(* Logix 5000 project; controller R400_500_XLS vendor 1 type 14 code 216 rev 31.11; software revision 31.01; part 16 of 32 *)
(* tags used below, declared in another part *)
   CycleModifBuffer : UDT_CYCLE;
   DRYING : DINT;   // Drying id number
   DRYING_HEAT_SENSITIVE_SEL : DINT;   // Drying heat sensitive
   DRYING_MODE_SEL : DINT;   // Drying mode selector index
   DRYING_TEMP_C_SEL : DINT;   // Drying temperature index
   DRYING_TEMP_F_SEL : DINT;   // Drying temperature index
   DRYING_TIME_MIN_NUM : DINT;   // Drying time (minutes) numeric input index
   DRYING_TIME_SEC_NUM : DINT;   // Drying time (seconds) numeric input index
   FC83_DryHeatSensitive : DINT;   // Drying is heat sensitive?
   FC83_DryTemp : DINT;   // Drying temperature (hi/low)
   FC83_FRinse_Drained : DINT;   // Drained final rinse flag
   FC83_FRinse_Heated : DINT;   // Heated final rinse flag
   FC83_FRinse_Recirculated : DINT;   // Recirculated final rinse flag
   FC83_ONS : SINT;
   FRINSE_COND_SET_POINT_NUM : DINT;   // Final rinse conductivity set point numeric input index
   FRINSE_DRAIN_SEL : DINT;   // Final rinse drained selector's index
   FRINSE_HEATING_SEL : DINT;   // Final rinse heating selector's index
   FRINSE_MIN_NUMBER_NUM : DINT;   // Final rinse minimum number of final rinse numeric input index
   FRINSE_NUMBER_NUM : DINT;   // Final rinse number of final rinse numeric input index
   FRINSE_RECIRC_SEL : DINT;   // Final rinse recirculated selector's index
   FRINSE_TIME_MIN_NUM : DINT;   // Final rinse time (minutes) numeric input index
   FRINSE_TIME_SEC_NUM : DINT;   // Final rinse time (seconds) numeric input index
   FRINSE_TYPE_SEL : DINT;   // Final rinse type selector's index
   M : DINT[5];   // Memory Bits
   MaxTrtTempSp : REAL;
   NON_RECIRCULATED_FINAL_RINSE_MINUTES : DINT;   // Number of minutes for the non recirculated final rinse
   NON_RECIRCULATED_FINAL_RINSE_SECONDS : DINT;   // Number of seconds for the non recirculated final rinse
   Rinse_Select : BOOL;
   RinseIndex : SINT;
   Second_Inj_conc : BOOL;
   WashIndex : SINT;
   cfgRinseHeated : SINT;
   cfgRinseMin : SINT;
   cfgRinseSec : SINT;
   CfgRinseTempSp : REAL;
   cfgRinseWport : SINT;
   CfgWshInjRateImperial : REAL;   // Wash Injection Rate - Oz / Gal
   CfgWshInjRateMetric : REAL;   // Wash Injection Rate - mL / L
   ChemConcUnit : BOOL;   // 0 = mL/L; 1 = oz/gal
   Msg_TempSp : SINT;   // HMI Information Message tag
   NumInput : UDT_NUMERIC_INPUT[65];   // Numeric input
   NumInputReal : UDT_NUMERIC_INPUT_REAL[17];
   Screen_Ctrl : DINT;   // PLC Screen Request
   Selector : UDT_SELECTOR[25];   // Piloted list selector
   TempUnit : BOOL;   // Temperature Units 0= Celcius 1 = Farhenheit
   Tpb : DINT[11];
   TpbImage : DINT[11];
   udtFRHeatingSel : UDT_SELECTOR;
   udtFRLastRinseDrained : UDT_SELECTOR;
   udtFRRecirculation : UDT_SELECTOR;
   udtFRType : UDT_SELECTOR;
   Unit : Hrdwre;   // Unit Configuration
(* MainProgram, continued *)

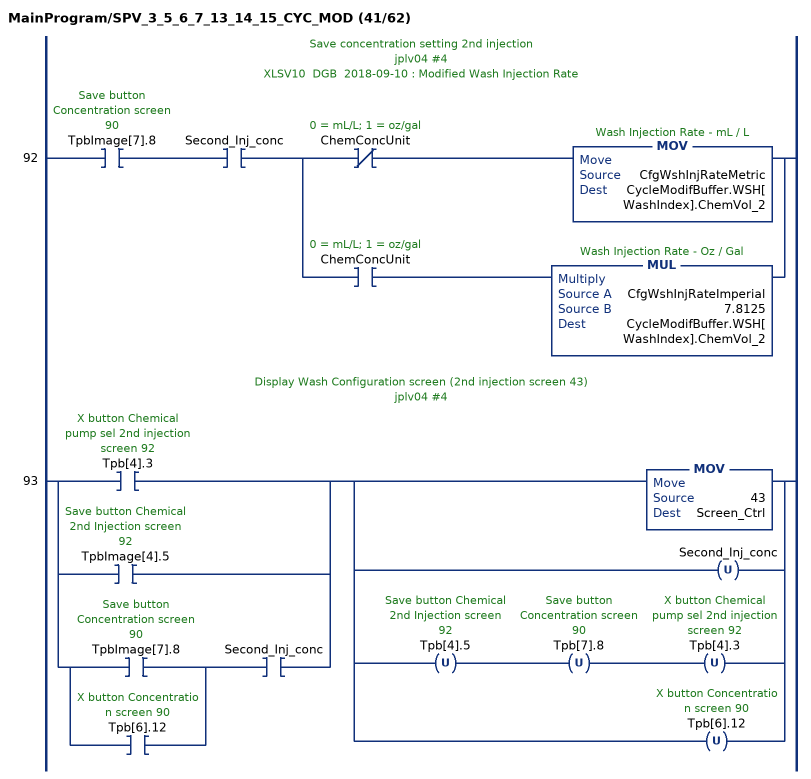
   [picture p292: MainProgram/SPV_3_5_6_7_13_14_15_CYC_MOD rungs 92-93]
   // Save concentration setting 2nd injection
   // jplv04 #4
   // XLSV10  DGB  2018-09-10 : Modified Wash Injection Rate
   92: XIC(TpbImage[7].8)XIC(Second_Inj_conc)[XIO(ChemConcUnit) MOV(CfgWshInjRateMetric,CycleModifBuffer.WSH[WashIndex].ChemVol_2) ,XIC(ChemConcUnit) MUL(CfgWshInjRateImperial,7.8125,CycleModifBuffer.WSH[WashIndex].ChemVol_2) ];
   // Display Wash Configuration screen (2nd injection screen 43)
   // jplv04 #4
   93: [XIC(Tpb[4].3) ,XIC(TpbImage[4].5) ,[XIC(TpbImage[7].8) ,XIC(Tpb[6].12) ] XIC(Second_Inj_conc) ][MOV(43,Screen_Ctrl) ,OTU(Second_Inj_conc) ,OTU(Tpb[4].5) OTU(Tpb[7].8) OTU(Tpb[4].3) ,OTU(Tpb[6].12) ];
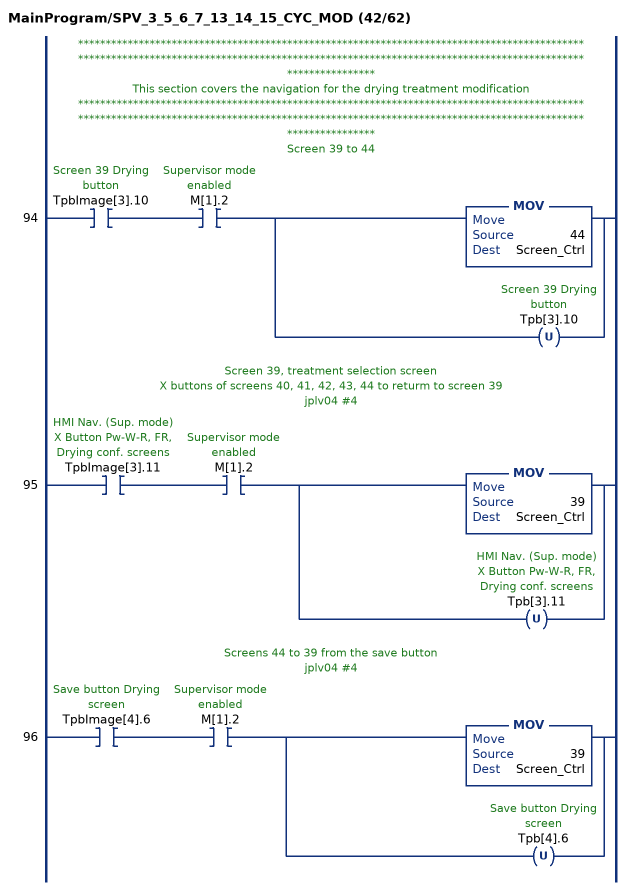
   // ********************************************************************************************************************************************************************************************************
   // This section covers the navigation for the drying treatment modification
   // ********************************************************************************************************************************************************************************************************
   // Screen 39 to 44
   94: XIC(TpbImage[3].10)XIC(M[1].2)[MOV(44,Screen_Ctrl) ,OTU(Tpb[3].10) ];
   // Screen 39, treatment selection screen
   // X buttons of screens 40, 41, 42, 43, 44 to returm to screen 39
   // jplv04 #4
   95: XIC(TpbImage[3].11)XIC(M[1].2)[MOV(39,Screen_Ctrl) ,OTU(Tpb[3].11) ];
   // Screens 44 to 39 from the save button
   // jplv04 #4
   96: XIC(TpbImage[4].6)XIC(M[1].2)[MOV(39,Screen_Ctrl) ,OTU(Tpb[4].6) ];
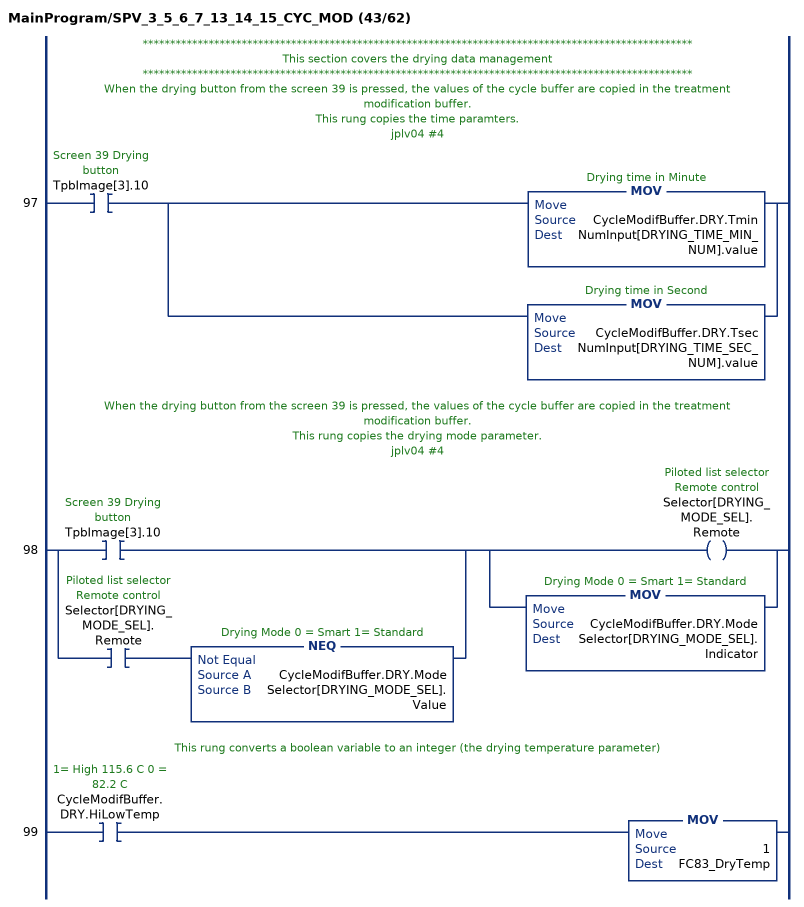
   // ****************************************************************************************************
   // This section covers the drying data management
   // ****************************************************************************************************
   // When the drying button from the screen 39 is pressed, the values of the cycle buffer are copied in the treatment modification buffer.
   // This rung copies the time paramters.
   // jplv04 #4
   97: XIC(TpbImage[3].10)[MOV(CycleModifBuffer.DRY.Tmin,NumInput[DRYING_TIME_MIN_NUM].value) ,MOV(CycleModifBuffer.DRY.Tsec,NumInput[DRYING_TIME_SEC_NUM].value) ];
   // When the drying button from the screen 39 is pressed, the values of the cycle buffer are copied in the treatment modification buffer.
   // This rung copies the drying mode parameter.
   // jplv04 #4
   98: [XIC(TpbImage[3].10) ,XIC(Selector[DRYING_MODE_SEL].Remote) NEQ(CycleModifBuffer.DRY.Mode,Selector[DRYING_MODE_SEL].Value) ][OTE(Selector[DRYING_MODE_SEL].Remote) ,MOV(CycleModifBuffer.DRY.Mode,Selector[DRYING_MODE_SEL].Indicator) ];
   // This rung converts a boolean variable to an integer (the drying temperature parameter)
   99: XIC(CycleModifBuffer.DRY.HiLowTemp)MOV(1,FC83_DryTemp);
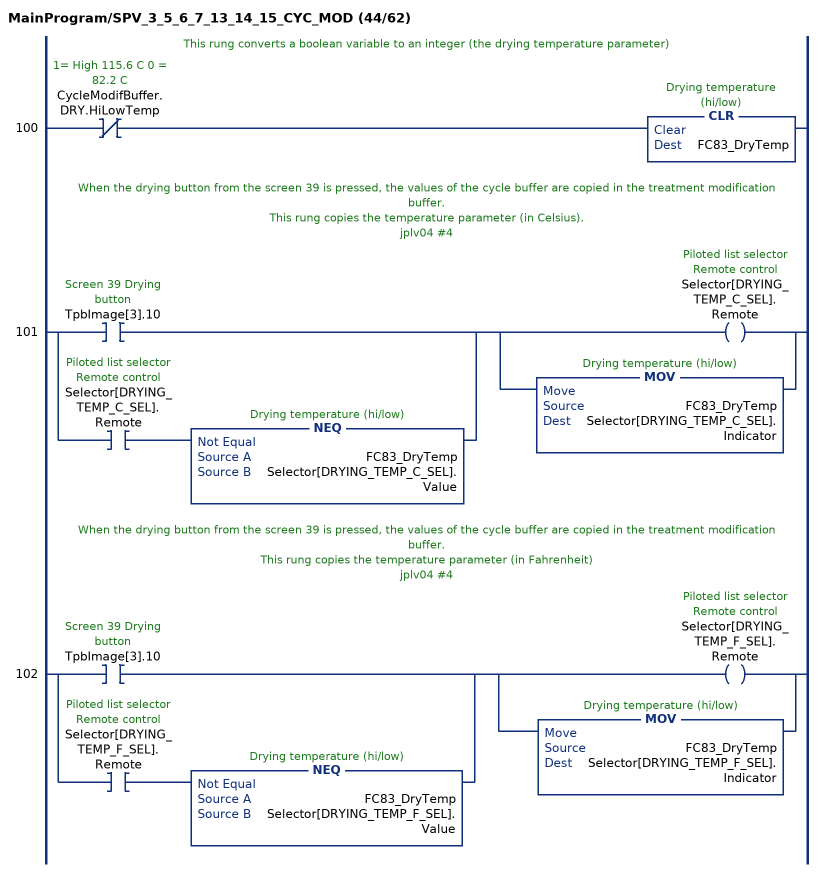
   // This rung converts a boolean variable to an integer (the drying temperature parameter)
   100: XIO(CycleModifBuffer.DRY.HiLowTemp)CLR(FC83_DryTemp);
   // When the drying button from the screen 39 is pressed, the values of the cycle buffer are copied in the treatment modification buffer.
   // This rung copies the temperature parameter (in Celsius).
   // jplv04 #4
   101: [XIC(TpbImage[3].10) ,XIC(Selector[DRYING_TEMP_C_SEL].Remote) NEQ(FC83_DryTemp,Selector[DRYING_TEMP_C_SEL].Value) ][OTE(Selector[DRYING_TEMP_C_SEL].Remote) ,MOV(FC83_DryTemp,Selector[DRYING_TEMP_C_SEL].Indicator) ];
   // When the drying button from the screen 39 is pressed, the values of the cycle buffer are copied in the treatment modification buffer.
   // This rung copies the temperature parameter (in Fahrenheit)
   // jplv04 #4
   102: [XIC(TpbImage[3].10) ,XIC(Selector[DRYING_TEMP_F_SEL].Remote) NEQ(FC83_DryTemp,Selector[DRYING_TEMP_F_SEL].Value) ][OTE(Selector[DRYING_TEMP_F_SEL].Remote) ,MOV(FC83_DryTemp,Selector[DRYING_TEMP_F_SEL].Indicator) ];
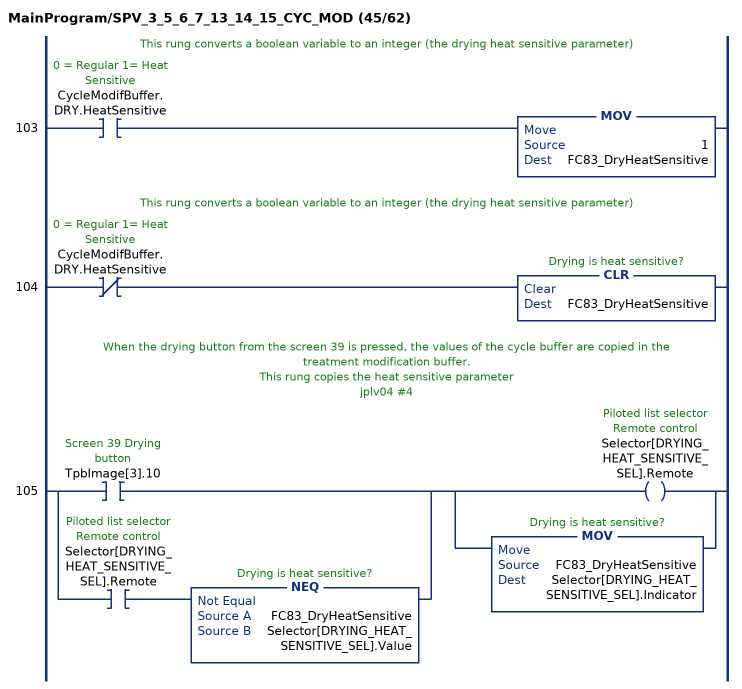
   // This rung converts a boolean variable to an integer (the drying heat sensitive parameter)
   103: XIC(CycleModifBuffer.DRY.HeatSensitive)MOV(1,FC83_DryHeatSensitive);
   // This rung converts a boolean variable to an integer (the drying heat sensitive parameter)
   104: XIO(CycleModifBuffer.DRY.HeatSensitive)CLR(FC83_DryHeatSensitive);
   // When the drying button from the screen 39 is pressed, the values of the cycle buffer are copied in the treatment modification buffer.
   // This rung copies the heat sensitive parameter
   // jplv04 #4
   105: [XIC(TpbImage[3].10) ,XIC(Selector[DRYING_HEAT_SENSITIVE_SEL].Remote) NEQ(FC83_DryHeatSensitive,Selector[DRYING_HEAT_SENSITIVE_SEL].Value) ][OTE(Selector[DRYING_HEAT_SENSITIVE_SEL].Remote) ,MOV(FC83_DryHeatSensitive,Selector[DRYING_HEAT_SENSITIVE_SEL].Indicator) ];
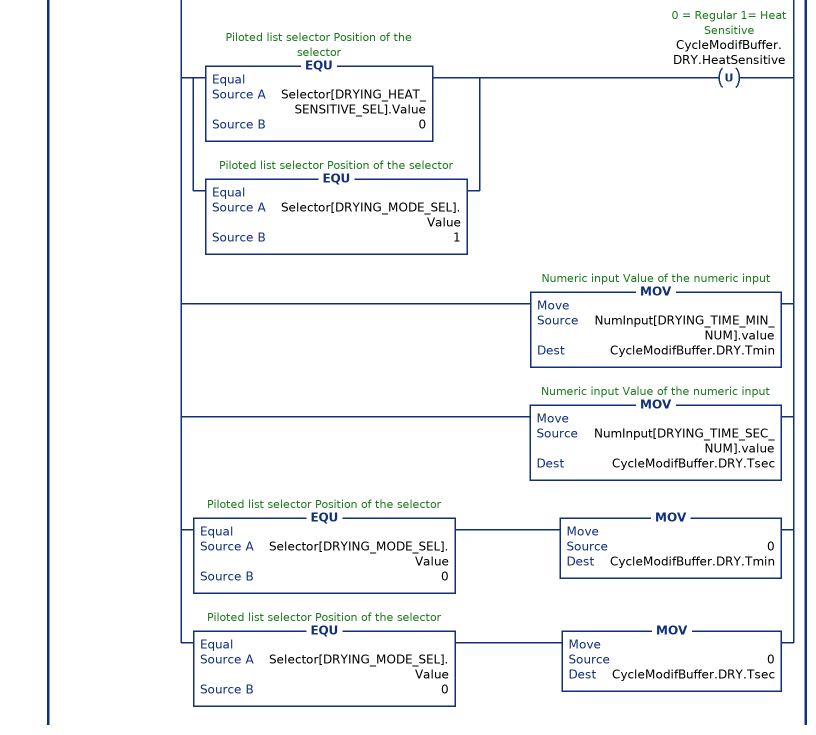
   // When the save button is pressed, the values are copied from the drying modification buffer to the cycle modification buffer
   // jplv04 #4
   106: XIC(TpbImage[4].6)[MOV(Selector[DRYING_MODE_SEL].Value,CycleModifBuffer.DRY.Mode) ,[XIO(TempUnit) EQU(Selector[DRYING_TEMP_C_SEL].Value,1) ,XIC(TempUnit) EQU(Selector[DRYING_TEMP_F_SEL].Value,1) ] OTL(CycleModifBuffer.DRY.HiLowTemp) ,[XIC(TempUnit) EQU(Selector[DRYING_TEMP_F_SEL].Value,0) ,XIO(TempUnit) EQU(Selector[DRYING_TEMP_C_SEL].Value,0) ,EQU(Selector[DRYING_MODE_SEL].Value,0) ] OTU(CycleModifBuffer.DRY.HiLowTemp) ,EQU(Selector[DRYING_HEAT_SENSITIVE_SEL].Value,1) OTL(CycleModifBuffer.DRY.HeatSensitive) ,[EQU(Selector[DRYING_HEAT_SENSITIVE_SEL].Value,0) ,EQU(Selector[DRYING_MODE_SEL].Value,1) ] OTU(CycleModifBuffer.DRY.HeatSensitive) ,MOV(NumInput[DRYING_TIME_MIN_NUM].value,CycleModifBuffer.DRY.Tmin) ,MOV(NumInput[DRYING_TIME_SEC_NUM].value,CycleModifBuffer.DRY.Tsec) ,EQU(Selector[DRYING_MODE_SEL].Value,0) MOV(0,CycleModifBuffer.DRY.Tmin) ,EQU(Selector[DRYING_MODE_SEL].Value,0) MOV(0,CycleModifBuffer.DRY.Tsec) ];
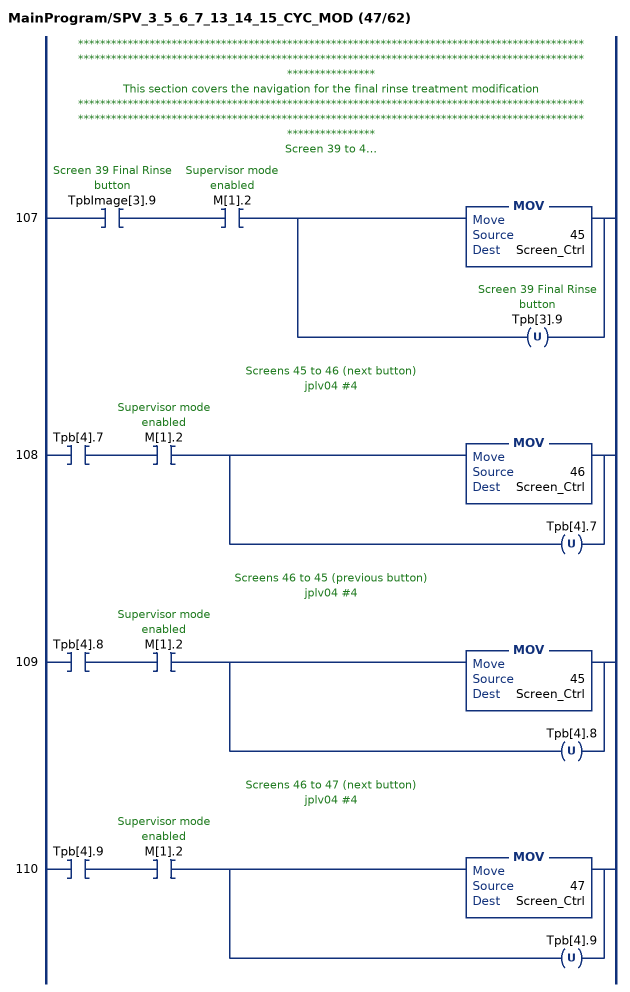
   // ********************************************************************************************************************************************************************************************************
   // This section covers the navigation for the final rinse treatment modification
   // ********************************************************************************************************************************************************************************************************
   // Screen 39 to 45
   // jplv04 #4
   107: XIC(TpbImage[3].9)XIC(M[1].2)[MOV(45,Screen_Ctrl) ,OTU(Tpb[3].9) ];
   // Screens 45 to 46 (next button)
   // jplv04 #4
   108: XIC(Tpb[4].7)XIC(M[1].2)[MOV(46,Screen_Ctrl) ,OTU(Tpb[4].7) ];
   // Screens 46 to 45 (previous button)
   // jplv04 #4
   109: XIC(Tpb[4].8)XIC(M[1].2)[MOV(45,Screen_Ctrl) ,OTU(Tpb[4].8) ];
   // Screens 46 to 47 (next button)
   // jplv04 #4
   110: XIC(Tpb[4].9)XIC(M[1].2)[MOV(47,Screen_Ctrl) ,OTU(Tpb[4].9) ];
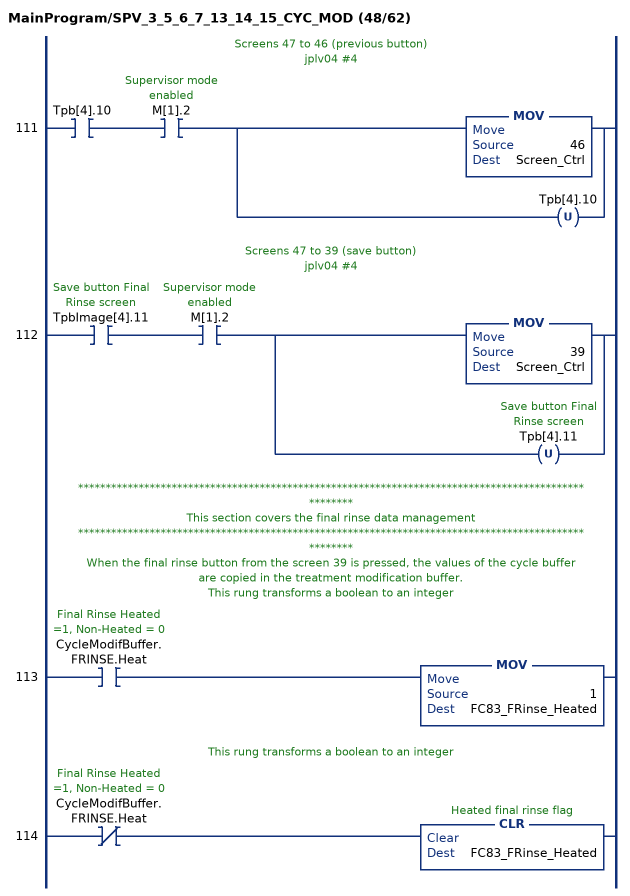
   // Screens 47 to 46 (previous button)
   // jplv04 #4
   111: XIC(Tpb[4].10)XIC(M[1].2)[MOV(46,Screen_Ctrl) ,OTU(Tpb[4].10) ];
   // Screens 47 to 39 (save button)
   // jplv04 #4
   112: XIC(TpbImage[4].11)XIC(M[1].2)[MOV(39,Screen_Ctrl) ,OTU(Tpb[4].11) ];
   // ****************************************************************************************************
   // This section covers the final rinse data management
   // ****************************************************************************************************
   // When the final rinse button from the screen 39 is pressed, the values of the cycle buffer are copied in the treatment modification buffer.
   // This rung transforms a boolean to an integer
   113: XIC(CycleModifBuffer.FRINSE.Heat)MOV(1,FC83_FRinse_Heated);
   // This rung transforms a boolean to an integer
   114: XIO(CycleModifBuffer.FRINSE.Heat)CLR(FC83_FRinse_Heated);
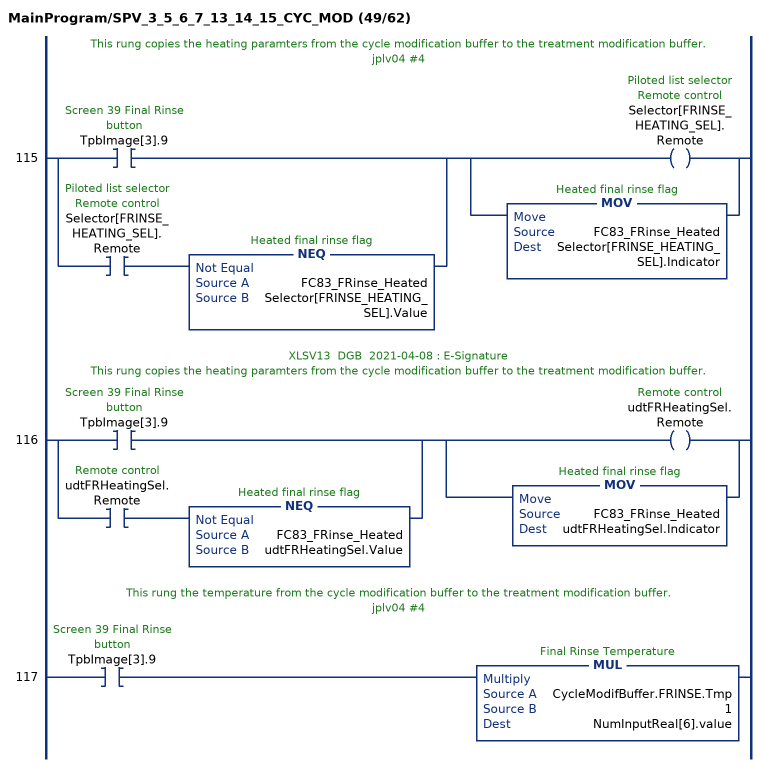
   // This rung copies the heating paramters from the cycle modification buffer to the treatment modification buffer.
   // jplv04 #4
   115: [XIC(TpbImage[3].9) ,XIC(Selector[FRINSE_HEATING_SEL].Remote) NEQ(FC83_FRinse_Heated,Selector[FRINSE_HEATING_SEL].Value) ][OTE(Selector[FRINSE_HEATING_SEL].Remote) ,MOV(FC83_FRinse_Heated,Selector[FRINSE_HEATING_SEL].Indicator) ];
   // XLSV13  DGB  2021-04-08 : E-Signature
   // This rung copies the heating paramters from the cycle modification buffer to the treatment modification buffer.
   116: [XIC(TpbImage[3].9) ,XIC(udtFRHeatingSel.Remote) NEQ(FC83_FRinse_Heated,udtFRHeatingSel.Value) ][OTE(udtFRHeatingSel.Remote) ,MOV(FC83_FRinse_Heated,udtFRHeatingSel.Indicator) ];
   // This rung the temperature from the cycle modification buffer to the treatment modification buffer.
   // jplv04 #4
   117: XIC(TpbImage[3].9)MUL(CycleModifBuffer.FRINSE.Tmp,1,NumInputReal[6].value);
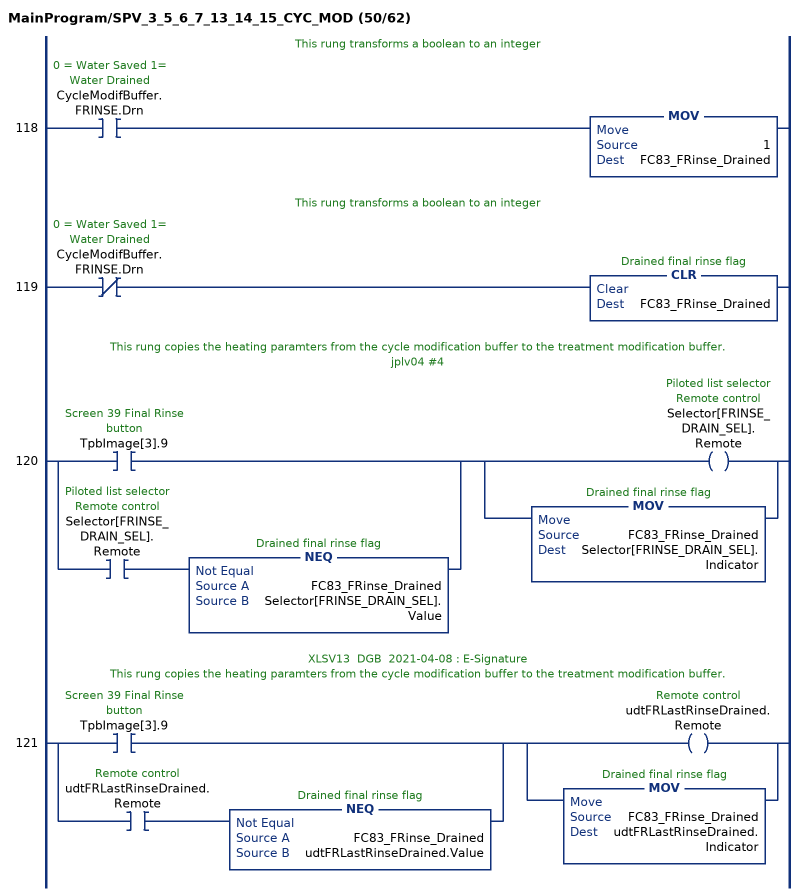
   // This rung transforms a boolean to an integer
   118: XIC(CycleModifBuffer.FRINSE.Drn)MOV(1,FC83_FRinse_Drained);
   // This rung transforms a boolean to an integer
   119: XIO(CycleModifBuffer.FRINSE.Drn)CLR(FC83_FRinse_Drained);
   // This rung copies the heating paramters from the cycle modification buffer to the treatment modification buffer.
   // jplv04 #4
   120: [XIC(TpbImage[3].9) ,XIC(Selector[FRINSE_DRAIN_SEL].Remote) NEQ(FC83_FRinse_Drained,Selector[FRINSE_DRAIN_SEL].Value) ][OTE(Selector[FRINSE_DRAIN_SEL].Remote) ,MOV(FC83_FRinse_Drained,Selector[FRINSE_DRAIN_SEL].Indicator) ];
   // XLSV13  DGB  2021-04-08 : E-Signature
   // This rung copies the heating paramters from the cycle modification buffer to the treatment modification buffer.
   121: [XIC(TpbImage[3].9) ,XIC(udtFRLastRinseDrained.Remote) NEQ(FC83_FRinse_Drained,udtFRLastRinseDrained.Value) ][OTE(udtFRLastRinseDrained.Remote) ,MOV(FC83_FRinse_Drained,udtFRLastRinseDrained.Indicator) ];
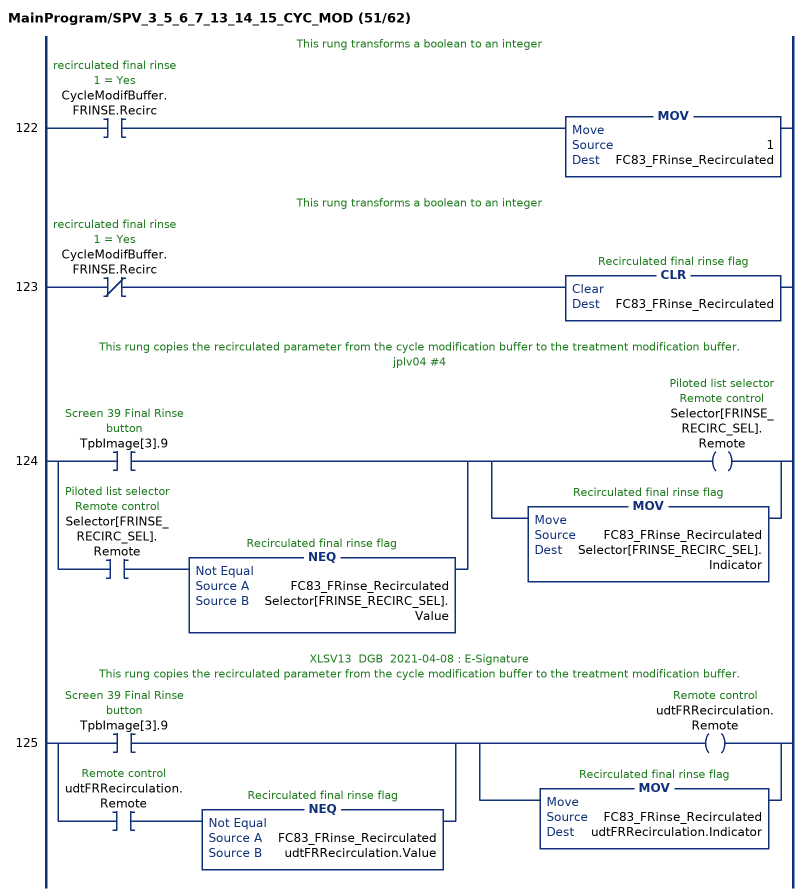
   // This rung transforms a boolean to an integer
   122: XIC(CycleModifBuffer.FRINSE.Recirc)MOV(1,FC83_FRinse_Recirculated);
   // This rung transforms a boolean to an integer
   123: XIO(CycleModifBuffer.FRINSE.Recirc)CLR(FC83_FRinse_Recirculated);
   // This rung copies the recirculated parameter from the cycle modification buffer to the treatment modification buffer.
   // jplv04 #4
   124: [XIC(TpbImage[3].9) ,XIC(Selector[FRINSE_RECIRC_SEL].Remote) NEQ(FC83_FRinse_Recirculated,Selector[FRINSE_RECIRC_SEL].Value) ][OTE(Selector[FRINSE_RECIRC_SEL].Remote) ,MOV(FC83_FRinse_Recirculated,Selector[FRINSE_RECIRC_SEL].Indicator) ];
   // XLSV13  DGB  2021-04-08 : E-Signature
   // This rung copies the recirculated parameter from the cycle modification buffer to the treatment modification buffer.
   125: [XIC(TpbImage[3].9) ,XIC(udtFRRecirculation.Remote) NEQ(FC83_FRinse_Recirculated,udtFRRecirculation.Value) ][OTE(udtFRRecirculation.Remote) ,MOV(FC83_FRinse_Recirculated,udtFRRecirculation.Indicator) ];
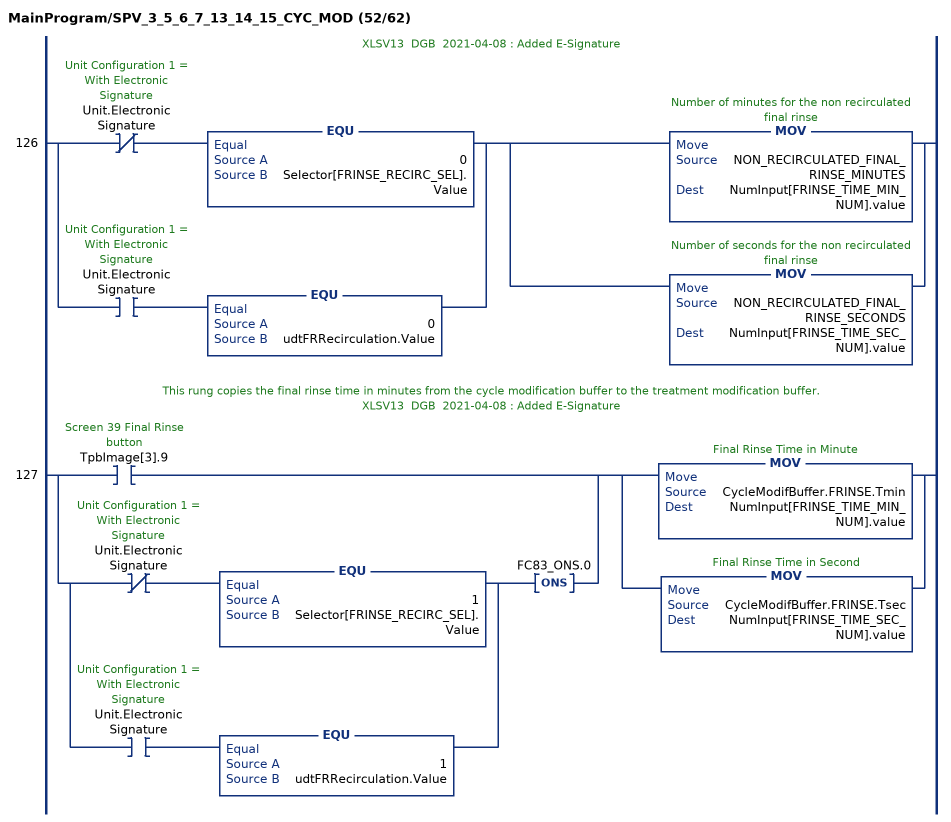
   // XLSV13  DGB  2021-04-08 : Added E-Signature
   126: [XIO(Unit.ElectronicSignature) EQU(0,Selector[FRINSE_RECIRC_SEL].Value) ,XIC(Unit.ElectronicSignature) EQU(0,udtFRRecirculation.Value) ][MOV(NON_RECIRCULATED_FINAL_RINSE_MINUTES,NumInput[FRINSE_TIME_MIN_NUM].value) ,MOV(NON_RECIRCULATED_FINAL_RINSE_SECONDS,NumInput[FRINSE_TIME_SEC_NUM].value) ];
   // This rung copies the final rinse time in minutes from the cycle modification buffer to the treatment modification buffer.
   // XLSV13  DGB  2021-04-08 : Added E-Signature
   127: [XIC(TpbImage[3].9) ,[XIO(Unit.ElectronicSignature) EQU(1,Selector[FRINSE_RECIRC_SEL].Value) ,XIC(Unit.ElectronicSignature) EQU(1,udtFRRecirculation.Value) ] ONS(FC83_ONS.0) ][MOV(CycleModifBuffer.FRINSE.Tmin,NumInput[FRINSE_TIME_MIN_NUM].value) ,MOV(CycleModifBuffer.FRINSE.Tsec,NumInput[FRINSE_TIME_SEC_NUM].value) ];
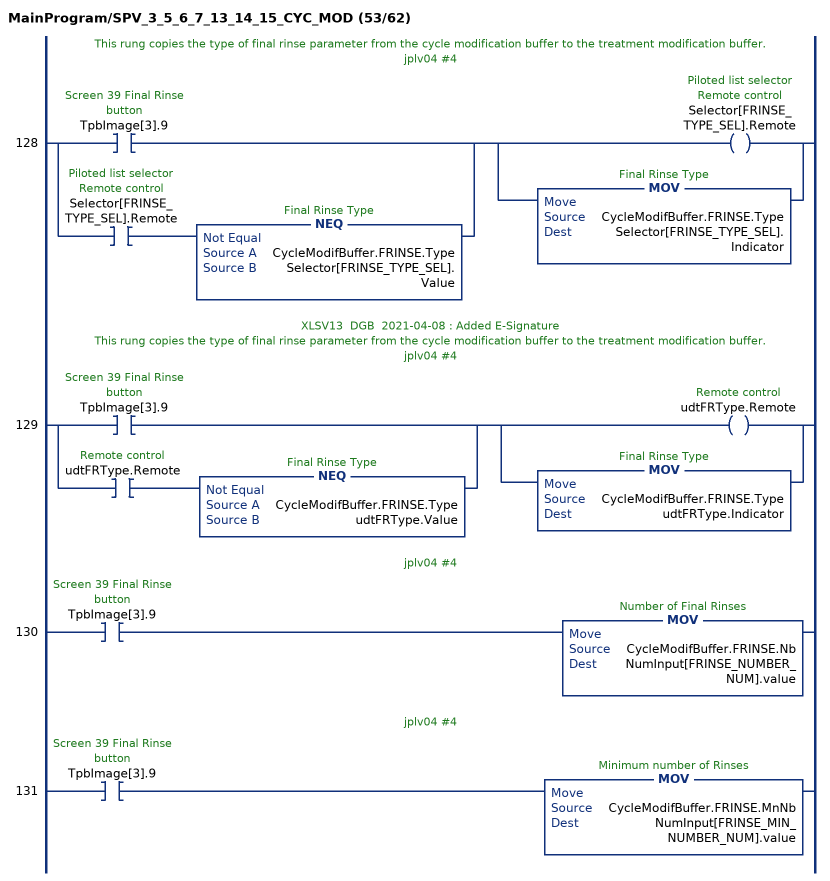
   // This rung copies the type of final rinse parameter from the cycle modification buffer to the treatment modification buffer.
   // jplv04 #4
   128: [XIC(TpbImage[3].9) ,XIC(Selector[FRINSE_TYPE_SEL].Remote) NEQ(CycleModifBuffer.FRINSE.Type,Selector[FRINSE_TYPE_SEL].Value) ][OTE(Selector[FRINSE_TYPE_SEL].Remote) ,MOV(CycleModifBuffer.FRINSE.Type,Selector[FRINSE_TYPE_SEL].Indicator) ];
   // XLSV13  DGB  2021-04-08 : Added E-Signature
   // This rung copies the type of final rinse parameter from the cycle modification buffer to the treatment modification buffer.
   // jplv04 #4
   129: [XIC(TpbImage[3].9) ,XIC(udtFRType.Remote) NEQ(CycleModifBuffer.FRINSE.Type,udtFRType.Value) ][OTE(udtFRType.Remote) ,MOV(CycleModifBuffer.FRINSE.Type,udtFRType.Indicator) ];
   // jplv04 #4
   130: XIC(TpbImage[3].9)MOV(CycleModifBuffer.FRINSE.Nb,NumInput[FRINSE_NUMBER_NUM].value);
   // jplv04 #4
   131: XIC(TpbImage[3].9)MOV(CycleModifBuffer.FRINSE.MnNb,NumInput[FRINSE_MIN_NUMBER_NUM].value);
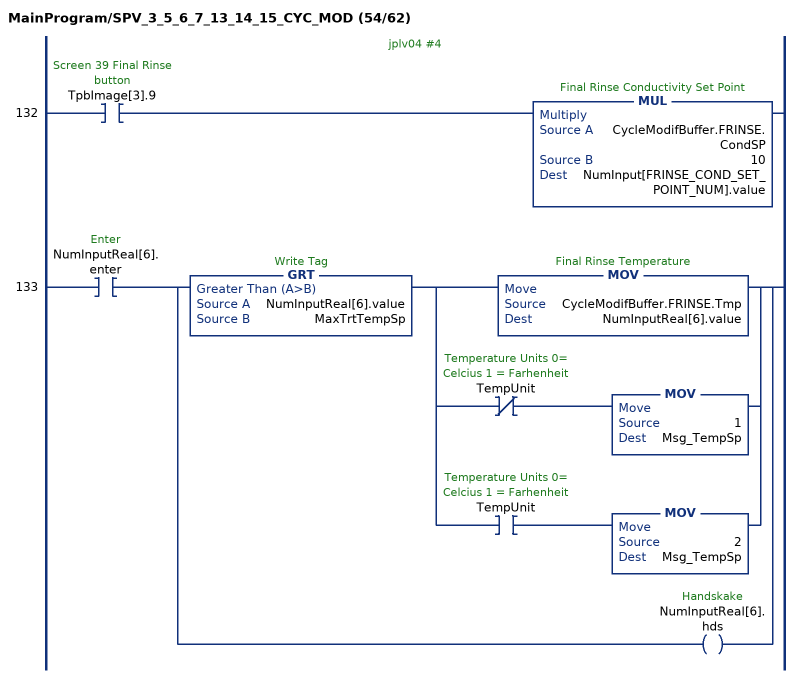
   // jplv04 #4
   132: XIC(TpbImage[3].9)MUL(CycleModifBuffer.FRINSE.CondSP,10,NumInput[FRINSE_COND_SET_POINT_NUM].value);
   133: XIC(NumInputReal[6].enter)[GRT(NumInputReal[6].value,MaxTrtTempSp) [MOV(CycleModifBuffer.FRINSE.Tmp,NumInputReal[6].value) ,XIO(TempUnit) MOV(1,Msg_TempSp) ,XIC(TempUnit) MOV(2,Msg_TempSp) ] ,OTE(NumInputReal[6].hds) ];
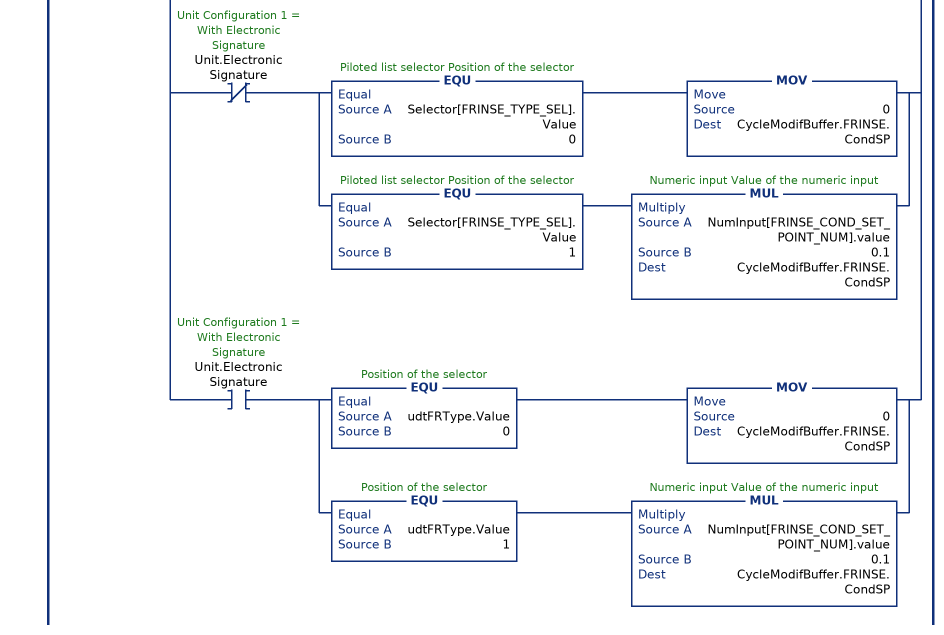
   // When the save button is pressed, the values are copied from the final rinse modification buffer to the cycle modification buffer
   // jplv04 #4
   // XLSV13  DGB  2021-04-08 : E-Signature
   134: XIC(TpbImage[4].11)[[XIO(Unit.ElectronicSignature) [EQU(Selector[FRINSE_HEATING_SEL].Value,1) OTL(CycleModifBuffer.FRINSE.Heat) ,EQU(Selector[FRINSE_HEATING_SEL].Value,0) OTU(CycleModifBuffer.FRINSE.Heat) ] ,XIC(Unit.ElectronicSignature) [EQU(udtFRHeatingSel.Value,1) OTL(CycleModifBuffer.FRINSE.Heat) ,EQU(udtFRHeatingSel.Value,0) OTU(CycleModifBuffer.FRINSE.Heat) ] ] ,[XIO(Unit.ElectronicSignature) [EQU(Selector[FRINSE_HEATING_SEL].Value,0) MOV(0,CycleModifBuffer.FRINSE.Tmp) ,EQU(Selector[FRINSE_HEATING_SEL].Value,1) MUL(NumInputReal[6].value,1,CycleModifBuffer.FRINSE.Tmp) ] ,XIC(Unit.ElectronicSignature) [EQU(udtFRHeatingSel.Value,0) MOV(0,CycleModifBuffer.FRINSE.Tmp) ,EQU(udtFRHeatingSel.Value,1) MUL(NumInputReal[6].value,1,CycleModifBuffer.FRINSE.Tmp) ] ] ,[XIO(Unit.ElectronicSignature) [EQU(Selector[FRINSE_DRAIN_SEL].Value,1) OTL(CycleModifBuffer.FRINSE.Drn) ,EQU(Selector[FRINSE_DRAIN_SEL].Value,0) OTU(CycleModifBuffer.FRINSE.Drn) ] ,XIC(Unit.ElectronicSignature) [EQU(udtFRLastRinseDrained.Value,1) OTL(CycleModifBuffer.FRINSE.Drn) ,EQU(udtFRLastRinseDrained.Value,0) OTU(CycleModifBuffer.FRINSE.Drn) ] ] ,[XIO(Unit.ElectronicSignature) [EQU(Selector[FRINSE_RECIRC_SEL].Value,1) OTL(CycleModifBuffer.FRINSE.Recirc) ,EQU(Selector[FRINSE_RECIRC_SEL].Value,0) OTU(CycleModifBuffer.FRINSE.Recirc) ] ,XIC(Unit.ElectronicSignature) [EQU(udtFRRecirculation.Value,1) OTL(CycleModifBuffer.FRINSE.Recirc) ,EQU(udtFRRecirculation.Value,0) OTU(CycleModifBuffer.FRINSE.Recirc) ] ] ,MOV(NumInput[FRINSE_TIME_MIN_NUM].value,CycleModifBuffer.FRINSE.Tmin) ,MOV(NumInput[FRINSE_TIME_SEC_NUM].value,CycleModifBuffer.FRINSE.Tsec) ,[XIO(Unit.ElectronicSignature) MOV(Selector[FRINSE_TYPE_SEL].Value,CycleModifBuffer.FRINSE.Type) ,XIC(Unit.ElectronicSignature) MOV(udtFRType.Value,CycleModifBuffer.FRINSE.Type) ] ,[XIO(Unit.ElectronicSignature) [EQU(Selector[FRINSE_TYPE_SEL].Value,0) MOV(NumInput[FRINSE_NUMBER_NUM].value,CycleModifBuffer.FRINSE.Nb) ,EQU(Selector[FRINSE_TYPE_SEL].Value,1) MOV(0,CycleModifBuffer.FRINSE.Nb) ] ,XIC(Unit.ElectronicSignature) [EQU(udtFRType.Value,0) MOV(NumInput[FRINSE_NUMBER_NUM].value,CycleModifBuffer.FRINSE.Nb) ,EQU(udtFRType.Value,1) MOV(0,CycleModifBuffer.FRINSE.Nb) ] ] ,[XIO(Unit.ElectronicSignature) [EQU(Selector[FRINSE_TYPE_SEL].Value,0) MOV(0,CycleModifBuffer.FRINSE.MnNb) ,EQU(Selector[FRINSE_TYPE_SEL].Value,1) MOV(NumInput[FRINSE_MIN_NUMBER_NUM].value,CycleModifBuffer.FRINSE.MnNb) ] ,XIC(Unit.ElectronicSignature) [EQU(udtFRType.Value,0) MOV(0,CycleModifBuffer.FRINSE.MnNb) ,EQU(udtFRType.Value,1) MOV(NumInput[FRINSE_MIN_NUMBER_NUM].value,CycleModifBuffer.FRINSE.MnNb) ] ] ,[XIO(Unit.ElectronicSignature) [EQU(Selector[FRINSE_TYPE_SEL].Value,0) MOV(0,CycleModifBuffer.FRINSE.CondSP) ,EQU(Selector[FRINSE_TYPE_SEL].Value,1) MUL(NumInput[FRINSE_COND_SET_POINT_NUM].value,0.1,CycleModifBuffer.FRINSE.CondSP) ] ,XIC(Unit.ElectronicSignature) [EQU(udtFRType.Value,0) MOV(0,CycleModifBuffer.FRINSE.CondSP) ,EQU(udtFRType.Value,1) MUL(NumInput[FRINSE_COND_SET_POINT_NUM].value,0.1,CycleModifBuffer.FRINSE.CondSP) ] ] ];
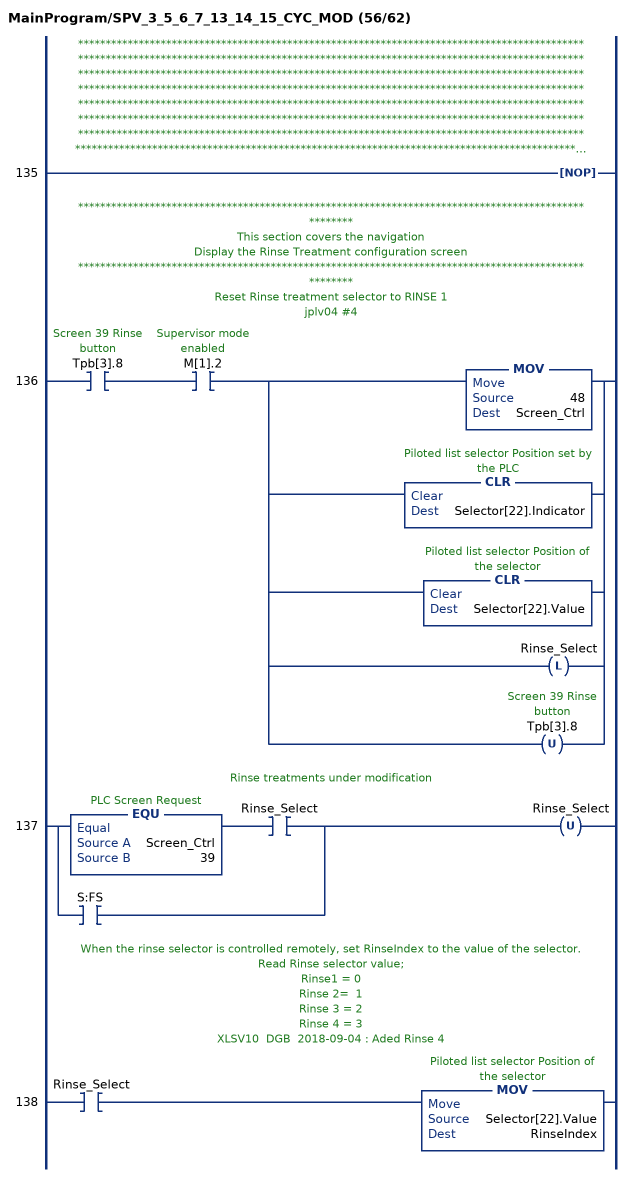
   // ****************************************************************************************************************************************************************************************************************************************************************************************************************************************************************************************************************************************************************************************************************************************************************************************************************************************************************************************************************************************************************************************************************************************************************************************************************************************************************************************************************************************************************************************************************************************************************************************************************************************************************************************************************************************************************************************************************************************************************************************************************************************************************************************************************************************************************************************************************************************************************************************************************************************************************************************************************************************************************************************************************************************************************************************************************************************************************************************************************************************************************************************************************************************************************************************
   135: NOP();
   // ****************************************************************************************************
   // This section covers the navigation
   // Display the Rinse Treatment configuration screen
   // ****************************************************************************************************
   // Reset Rinse treatment selector to RINSE 1
   // jplv04 #4
   136: XIC(Tpb[3].8)XIC(M[1].2)[MOV(48,Screen_Ctrl) ,CLR(Selector[22].Indicator) ,CLR(Selector[22].Value) ,OTL(Rinse_Select) ,OTU(Tpb[3].8) ];
   // Rinse treatments under modification
   137: [EQU(Screen_Ctrl,39) XIC(Rinse_Select) ,XIC(S:FS) ]OTU(Rinse_Select);
   // When the rinse selector is controlled remotely, set RinseIndex to the value of the selector.
   // Read Rinse selector value;
   // Rinse1 = 0
   // Rinse 2=  1
   // Rinse 3 = 2
   // Rinse 4 = 3
   // XLSV10  DGB  2018-09-04 : Aded Rinse 4
   138: XIC(Rinse_Select)MOV(Selector[22].Value,RinseIndex);
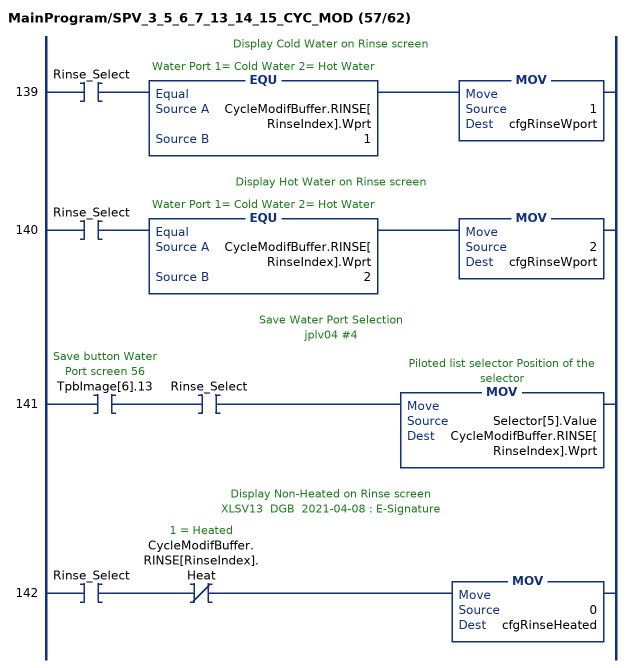
   // Display Cold Water on Rinse screen
   139: XIC(Rinse_Select)EQU(CycleModifBuffer.RINSE[RinseIndex].Wprt,1)MOV(1,cfgRinseWport);
   // Display Hot Water on Rinse screen
   140: XIC(Rinse_Select)EQU(CycleModifBuffer.RINSE[RinseIndex].Wprt,2)MOV(2,cfgRinseWport);
   // Save Water Port Selection
   // jplv04 #4
   141: XIC(TpbImage[6].13)XIC(Rinse_Select)MOV(Selector[5].Value,CycleModifBuffer.RINSE[RinseIndex].Wprt);
   // Display Non-Heated on Rinse screen
   // XLSV13  DGB  2021-04-08 : E-Signature
   142: XIC(Rinse_Select)XIO(CycleModifBuffer.RINSE[RinseIndex].Heat)MOV(0,cfgRinseHeated);
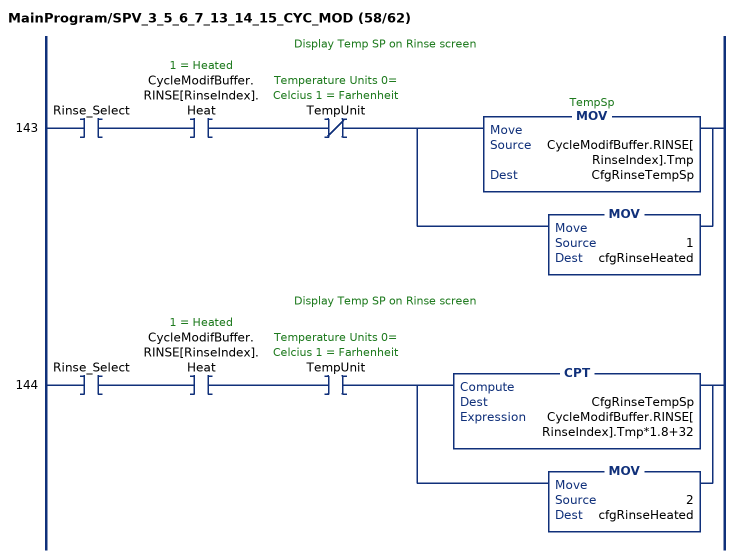
   // Display Temp SP on Rinse screen
   143: XIC(Rinse_Select)XIC(CycleModifBuffer.RINSE[RinseIndex].Heat)XIO(TempUnit)[MOV(CycleModifBuffer.RINSE[RinseIndex].Tmp,CfgRinseTempSp) ,MOV(1,cfgRinseHeated) ];
   // Display Temp SP on Rinse screen
   144: XIC(Rinse_Select)XIC(CycleModifBuffer.RINSE[RinseIndex].Heat)XIC(TempUnit)[CPT(CfgRinseTempSp,CycleModifBuffer.RINSE[RinseIndex].Tmp*1.8+32) ,MOV(2,cfgRinseHeated) ];
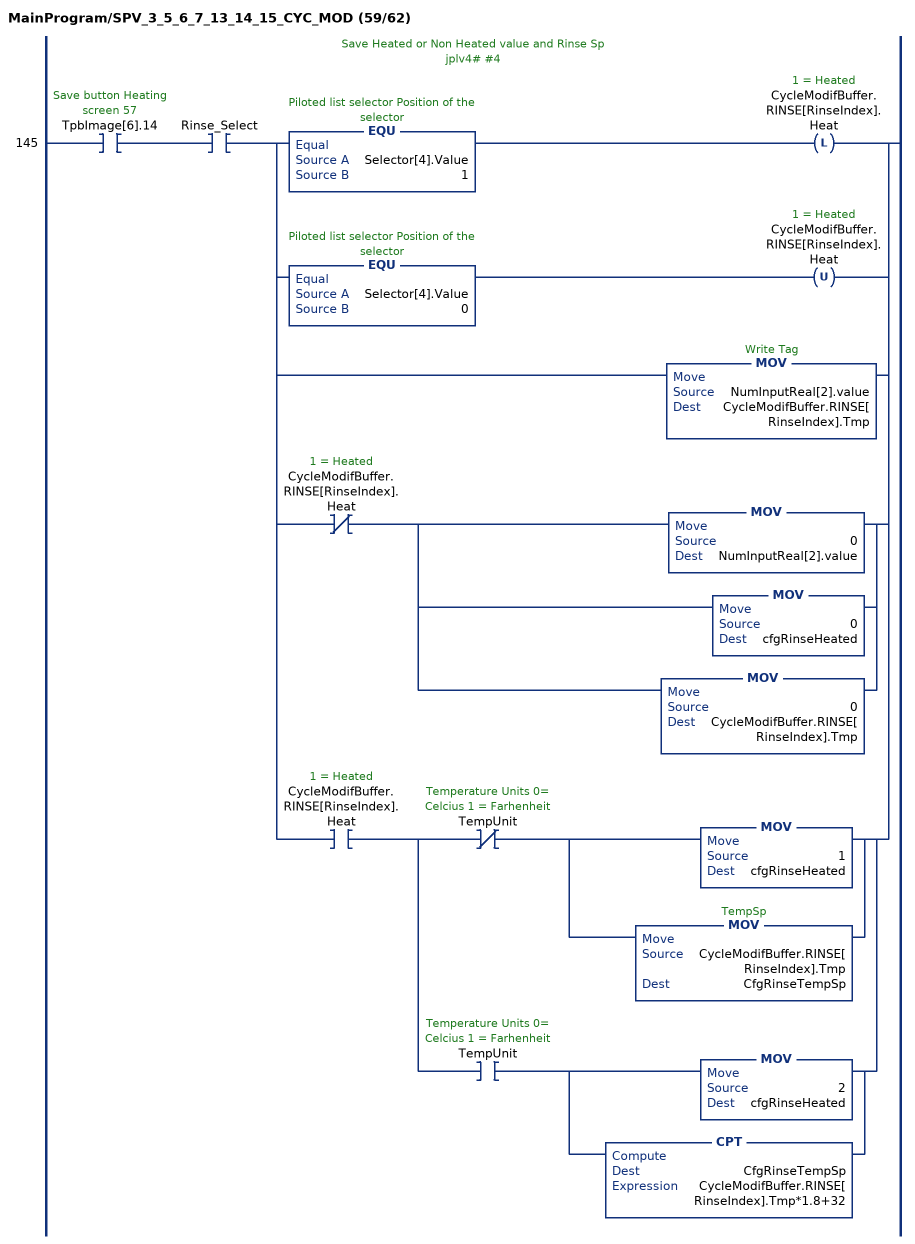
   // Save Heated or Non Heated value and Rinse Sp
   // jplv4# #4
   145: XIC(TpbImage[6].14)XIC(Rinse_Select)[EQU(Selector[4].Value,1) OTL(CycleModifBuffer.RINSE[RinseIndex].Heat) ,EQU(Selector[4].Value,0) OTU(CycleModifBuffer.RINSE[RinseIndex].Heat) ,MOV(NumInputReal[2].value,CycleModifBuffer.RINSE[RinseIndex].Tmp) ,XIO(CycleModifBuffer.RINSE[RinseIndex].Heat) [MOV(0,NumInputReal[2].value) ,MOV(0,cfgRinseHeated) ,MOV(0,CycleModifBuffer.RINSE[RinseIndex].Tmp) ] ,XIC(CycleModifBuffer.RINSE[RinseIndex].Heat) [XIO(TempUnit) [MOV(1,cfgRinseHeated) ,MOV(CycleModifBuffer.RINSE[RinseIndex].Tmp,CfgRinseTempSp) ] ,XIC(TempUnit) [MOV(2,cfgRinseHeated) ,CPT(CfgRinseTempSp,CycleModifBuffer.RINSE[RinseIndex].Tmp*1.8+32) ] ] ];
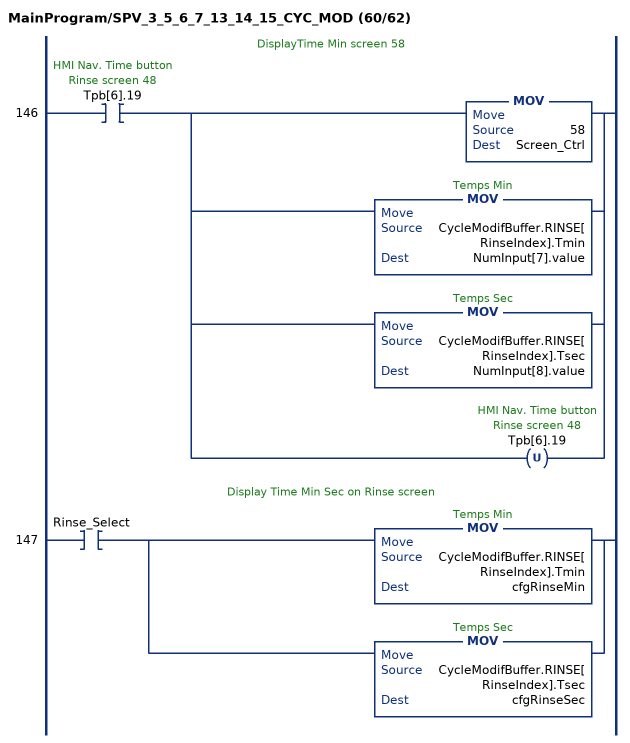
   // DisplayTime Min screen 58
   146: XIC(Tpb[6].19)[MOV(58,Screen_Ctrl) ,MOV(CycleModifBuffer.RINSE[RinseIndex].Tmin,NumInput[7].value) ,MOV(CycleModifBuffer.RINSE[RinseIndex].Tsec,NumInput[8].value) ,OTU(Tpb[6].19) ];
   // Display Time Min Sec on Rinse screen
   147: XIC(Rinse_Select)[MOV(CycleModifBuffer.RINSE[RinseIndex].Tmin,cfgRinseMin) ,MOV(CycleModifBuffer.RINSE[RinseIndex].Tsec,cfgRinseSec) ];
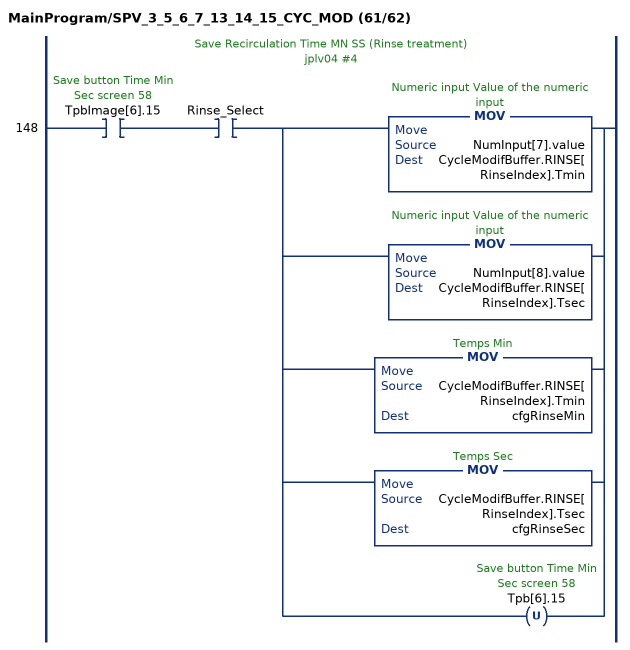
   // Save Recirculation Time MN SS (Rinse treatment)
   // jplv04 #4
   148: XIC(TpbImage[6].15)XIC(Rinse_Select)[MOV(NumInput[7].value,CycleModifBuffer.RINSE[RinseIndex].Tmin) ,MOV(NumInput[8].value,CycleModifBuffer.RINSE[RinseIndex].Tsec) ,MOV(CycleModifBuffer.RINSE[RinseIndex].Tmin,cfgRinseMin) ,MOV(CycleModifBuffer.RINSE[RinseIndex].Tsec,cfgRinseSec) ,OTU(Tpb[6].15) ];
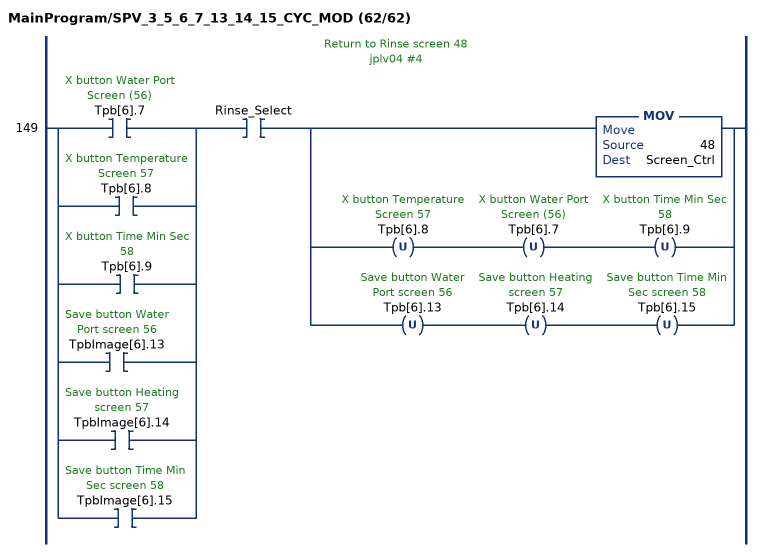
   // Return to Rinse screen 48
   // jplv04 #4
   149: [XIC(Tpb[6].7) ,XIC(Tpb[6].8) ,XIC(Tpb[6].9) ,XIC(TpbImage[6].13) ,XIC(TpbImage[6].14) ,XIC(TpbImage[6].15) ]XIC(Rinse_Select)[MOV(48,Screen_Ctrl) ,OTU(Tpb[6].8) OTU(Tpb[6].7) OTU(Tpb[6].9) ,OTU(Tpb[6].13) OTU(Tpb[6].14) OTU(Tpb[6].15) ];
END_ROUTINE
